(* IEC 61131-3 sources: axsharp/src/tests.integrations/integrated/src/ax/src/issues, 1 file *)

(* ---- GH_ISSUE_183.st ---- *)
NAMESPACE GH_ISSUE_183
    {S7.extern=ReadWrite}
    CLASS GH_ISSUE_183_1
        VAR PUBLIC
            NonZeroBasedArray : ARRAY[10..30] OF BYTE;
        END_VAR
    END_CLASS
END_NAMESPACE
